Fanuc KAREL source: KO00127.KL

PROGRAM KO00127
%NOLOCKGROUP
VAR
  A: ARRAY[2] OF SHORT
  B: ARRAY[2] OF SHORT
  OUT: INTEGER
BEGIN
  A[1] = 1
  B[1] = 2
  OUT = ATAN2(A[1], B[1])
END KO00127
